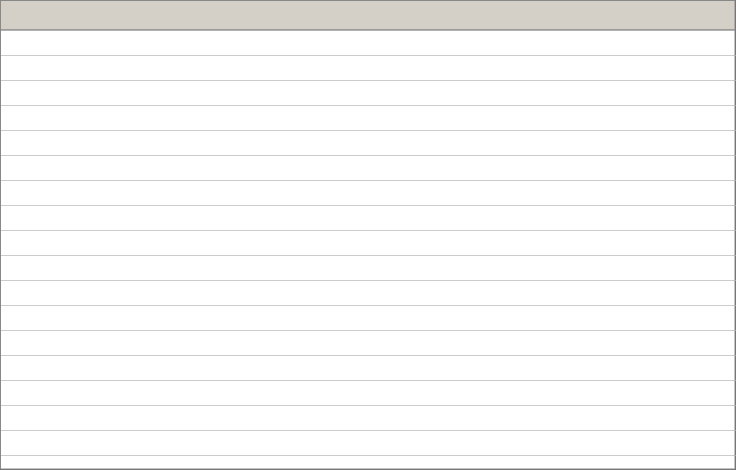
VISUALIZATION vis_Piston_Setting_Table  // 736x470
    Table (0,0 736x470), data array: stPisSetting
        p3854506369: stPisSetting[INDEX].t_minOpen
        p1892666644: stPisSetting[INDEX].t_minClose
        p338671338: stPisSetting[INDEX].t_maxOpen
        p2170511999: stPisSetting[INDEX].t_maxClose
        p3723444502: stPisSetting[INDEX].t_DelayOpen
        p1218418051: stPisSetting[INDEX].t_DelayClose
        p746581629: stPisSetting[INDEX].sen_Open_Exist
        p3104783080: stPisSetting[INDEX].sen_Close_Exist
END_VISUALIZATION

(* stored: Version 1.1.0.1, ProductVersion 3.1.4024.13
   Visu vis_Piston_Setting_Table: Id {96d7fd97-fcb8-471e-83e4-fa0e2d4fa8f3} *)
